{attribute 'qualified_only'}
{attribute 'strict'}
TYPE OUTPUT_ENUM :
(
	MONOSTABLE := 0,
	BISTABLE := 1
);
END_TYPE

(* stored: Version 1.1.0.1, ProductVersion 3.1.4024.12
   DUT OUTPUT_ENUM: Id {fd733a9e-f92f-442a-88d4-fb95da679b0a} *)
